FUNCTION_BLOCK FB_LogRecordProcessor_Mixin

PROPERTY pSelf : PVOID
GET
pSelf := THIS;
END_GET
END_PROPERTY

END_FUNCTION_BLOCK

(* stored: Version 1.1.0.1
   POU FB_LogRecordProcessor_Mixin: Id {3481a824-781e-4aa9-819e-1deb6d8b1261}, SpecialFunc None
   Property pSelf: Id {7e6151dd-6198-4fe1-9516-a1dfd6d8bdbe}
   Get Get: Id {7f117015-c51a-4865-8ea3-368656695039} *)
